INTERFACE I_Accelerometer

PROPERTY AccelerationInMPerS2 : Vector3
GET
END_GET
END_PROPERTY

PROPERTY TimestampInNs : ULINT
GET
END_GET
END_PROPERTY

PROPERTY IsValid : BOOL
GET
END_GET
END_PROPERTY

END_INTERFACE

(* stored: Version 1.1.0.1, ProductVersion 3.1.4026.12
   Itf I_Accelerometer: Id {4df7a45b-ba0b-5932-a8e0-8f729a3a027e}
   Property AccelerationInMPerS2: Id {38226d2c-778e-55a7-a7e6-c8884d8b7a30}
   Get Get: Id {4e4c0415-e88e-54aa-9f91-3b54d30c66b8}
   Property TimestampInNs: Id {33cf4371-98ef-5903-87e1-65261f5c03dd}
   Get Get: Id {857d7dca-706d-5711-af7d-94e17549a80c}
   Property IsValid: Id {2d77484d-cff3-5ede-86fe-65dc71906384}
   Get Get: Id {110d3938-ce3d-5afe-adbf-60330f7ba0d7} *)
